{attribute 'qualified_only'}
VAR_GLOBAL
	dwMicroSwitchDriverA AT %I* : DWORD;
	dwMicroSwitchDriverB AT %I* : DWORD;
END_VAR

(* stored: Version 1.1.0.1, ProductVersion 3.1.4024.15
   GVL GVL_MicroSwitch: Id {23487114-5e9f-4e40-92ef-271345d84160} *)
